(* PLC project g_tp_pulse, Anonymous Benchmark Suite 1.0 *)
(* stored: creationDateTime 2026-08-26T00:00:00 *)

PROGRAM g_tp_pulse
  VAR_INPUT
    Trig : BOOL;
  END_VAR
  VAR_OUTPUT
    Out : BOOL;
  END_VAR
  VAR
    TP0 : TP;
  END_VAR

(* LD diagram, written out as Structured Text *)
TP0(IN := Trig, PT := T#30ms);
Out := TP0.Q;
END_PROGRAM

CONFIGURATION Config0
  RESOURCE Res0 ON PLC
    TASK tcyclic(INTERVAL := T#10ms, PRIORITY := 0);
    PROGRAM inst0 WITH tcyclic : g_tp_pulse;
  END_RESOURCE
END_CONFIGURATION
